Staubli VAL3: program.dtx

mdesc mNomSpeed
bool bError
public num nLastIndex
